Fanuc KAREL source: KT00820.KL

PROGRAM KT00820
%NOLOCKGROUP
VAR
  I1: INTEGER
  I2: INTEGER
  OUT: INTEGER
BEGIN
  I1 = 2
  I2 = 3
  I1 = 2
  I2 = 3
  OUT = SIN(I1)
END KT00820
